TYPE ST_Safety_Speps :
STRUCT
	step1: BOOL;
	step2: BOOL;
	step3: BOOL;
	step4: BOOL;
	step5: BOOL;
	step6: BOOL;
	stepRnD	:	BOOL	;

END_STRUCT
END_TYPE

(* stored: Version 1.1.0.1, ProductVersion 3.1.4026.18
   DUT ST_Safety_Speps: Id {1b50b5e5-b749-4b15-b1ce-07d047ad7987} *)
